Fanuc KAREL source: ko00100.KL

PROGRAM KO00100
%STACKSIZE=65535
%PRIORITY=65535
%NOLOCKGROUP
VAR
A : INTEGER
B : REAL
OUT : REAL
BEGIN
A=1
B=2
-- UNRESOLVED_PC line 10 opcodes [27 27 21 64 22 76 23] marker_code=29
END KO00100
